// TIA Portal V20 export
// export: Created 2026-10-20T18:55:09.3234588Z, ExportSetting None, DisplayName Totally Integrated Automation Portal, DisplayVersion V20 Update 6, DisplayName TIA Portal Openness, DisplayVersion V20 Update 6, DisplayName TIA Portal Version Control Interface, DisplayVersion V20 Update 6, DisplayName SINAMICS Startdrive Advanced, DisplayVersion V20 SP1, DisplayName SINAMICS Startdrive G130, G150, S120, S150, SINAMICS MV, G220, S200, S210, DisplayVersion V20 SP1, DisplayName SINAMICS Startdrive G110M, G120, G120C, G120D, G120P, G115D, DisplayVersion V20 SP1, DisplayName STEP 7 Professional, DisplayVersion V20 Update 6, DisplayName STEP 7 Safety, DisplayVersion V20 Update 2, DisplayName WinCC Basic/Comfort/Advanced, DisplayVersion V20 Update 6, DisplayName WinCC Unified, DisplayVersion V20 Update 6
VAR_GLOBAL   // PLC tag table "IO_ET200_3"
   "C3204 - SENSOR CNV RIGHT (PALLET DETECT 1)" AT %I872.4 : Bool;
   "C3205 - SENSOR CNV RIGHT (PALLET DETECT 1)" AT %I874.4 : Bool;
   "C3207 - SENSOR CNV RIGHT (PALLET DETECT 1)" AT %I878.4 : Bool;
   "E-STOP L1 - CH1(3)" AT %I1662.0 : Bool;
   "E-STOP L2 - CH1(3)" AT %I1662.2 : Bool;
   "KEY REMOTE/LOCAL L1 - CH1(3)" AT %I1662.1 : Bool;
   "KEY REMOTE/LOCAL L2 - CH1(3)" AT %I1662.3 : Bool;
   "E-STOP L1 - CH2(3)" AT %I1662.4 : Bool;
   "KEY REMOTE/LOCAL L1 - CH2(3)" AT %I1662.5 : Bool;
   "E-STOP L2 - CH2(3)" AT %I1662.6 : Bool;
   "KEY REMOTE/LOCAL L2 - CH2(3)" AT %I1662.7 : Bool;
   "E-STOP L3 - CH1(3)" AT %I1670.0 : Bool;
   "KEY REMOTE/LOCAL L3 - CH1(3)" AT %I1670.1 : Bool;
   "E-STOP L4 - CH1(3)" AT %I1670.2 : Bool;
   "KEY REMOTE/LOCAL L4 - CH1(3)" AT %I1670.3 : Bool;
   "E-STOP L3 - CH2(3)" AT %I1670.4 : Bool;
   "KEY REMOTE/LOCAL L3 - CH2(3)" AT %I1670.5 : Bool;
   "E-STOP L4 - CH2(3)" AT %I1670.6 : Bool;
   "KEY REMOTE/LOCAL L4 - CH2(3)" AT %I1670.7 : Bool;
   "E-STOP L5 - CH1(3)" AT %I1678.0 : Bool;
   "KEY REMOTE/LOCAL L5 - CH1(3)" AT %I1678.1 : Bool;
   "E-STOP L6 - CH1(3)" AT %I1678.2 : Bool;
   "KEY REMOTE/LOCAL L6 - CH1(3)" AT %I1678.3 : Bool;
   "E-STOP L5 - CH2(3)" AT %I1678.4 : Bool;
   "KEY REMOTE/LOCAL L5 - CH2(3)" AT %I1678.5 : Bool;
   "E-STOP L6 - CH2(3)" AT %I1678.6 : Bool;
   "KEY REMOTE/LOCAL L6 - CH2(3)" AT %I1678.7 : Bool;
   "E-STOP L8 - CH1(3)" AT %I1686.2 : Bool;
   "KEY REMOTE/LOCAL L8 - CH1(3)" AT %I1686.3 : Bool;
   "E-STOP L8 - CH2(3)" AT %I1686.6 : Bool;
   "KEY REMOTE/LOCAL L8 - CH2(3)" AT %I1686.7 : Bool;
   "C3201 - SENSOR CNV RIGHT (PALLET DETECT 1)" AT %I866.4 : Bool;
   "C3201 - SHUTTLE IN POSITION 2" AT %I867.6 : Bool;
   "CVTD3 SENSOR CONVEYOR LEFT (PALLET DETECT 1)" AT %I140.2 : Bool;
   "C3201 - SENSOR CNV RIGHT (PALLET DETECT 2)" AT %I867.1 : Bool;
   "VTD3 DOCKING PINS EXTENDED 1" AT %I141.0 : Bool;
   "VTD3 LEVEL DETECT 1" AT %I141.7 : Bool;
   "C3201 - SENSOR CNV LEFT (FWD)" AT %I867.4 : Bool;
   "VTD3 DOCKING PINS EXTENDED 2" AT %I141.2 : Bool;
   "VTD3 LEVEL DETECT 2" AT %I141.6 : Bool;
   "C3201 - SHUTTLE IN POSITION 1" AT %I867.7 : Bool;
   "VTD3 DOCKING PINS RETRACTED 1" AT %I141.1 : Bool;
   "CVTD3 SENSOR CONVEYOR CENTER" AT %I140.3 : Bool;
   "VTD3 ULTIMATE SLOWDOWN" AT %I141.4 : Bool;
   "VTD3 ULTIMATE CREEP" AT %I141.5 : Bool;
   "CVTD3 SENSOR CONVEYOR RIGHT (PALLET DETECT 1)" AT %I140.5 : Bool;
   "CVTD3 SENSOR CONVEYOR LEFT (FWD)" AT %I140.1 : Bool;
   "VTD3 DOCKING PINS RETRACTED 2" AT %I141.3 : Bool;
   "C3201 - SENSOR CNV RIGHT (BWD)" AT %I866.5 : Bool;
   "C3201 - SENSOR CNV LEFT (PALLET DETECT 2)" AT %I867.0 : Bool;
   "C3201 - SENSOR CNV LEFT (PALLET DETECT 1)" AT %I867.5 : Bool;
   "CVTD3 SENSOR CONVEYOR RIGHT (BWD)" AT %I140.4 : Bool;
   "C3106 - SENSOR CNV RIGHT (PALLET DETECT 1)" AT %I861.5 : Bool;
   "C3208 - SENSOR CNV LEFT (FWD)" AT %I881.4 : Bool;
   "C3108 - SENSOR CNV LEFT (FWD)" AT %I864.5 : Bool;
   "C3107 - SENSOR CNV LEFT (PALLET DETECT 1)" AT %I862.4 : Bool;
   "C3107 - SENSOR CNV RIGHT (PALLET DETECT 2)" AT %I863.0 : Bool;
   "C3107 - SENSOR SAFETY PIN1 DOWN" AT %I863.3 : Bool;
   "C3208 - SENSOR SAFETY PIN1 UP" AT %I881.2 : Bool;
   "C3208 - SENSOR SAFETY PIN1 DOWN" AT %I881.3 : Bool;
   "C3108 - SENSOR SAFETY PIN1 DOWN" AT %I865.3 : Bool;
   "C3108 - SENSOR CNV RIGHT (PALLET DETECT 1)" AT %I865.5 : Bool;
   "C3207 - SENSOR CNV LEFT (PALLET DETECT 1)" AT %I879.1 : Bool;
   "C3106 - SENSOR SAFETY PIN1 DOWN" AT %I861.3 : Bool;
   "C3207 - SENSOR CNV RIGHT (PALLET DETECT 2)" AT %I879.5 : Bool;
   "C3106 - SENSOR CNV LEFT (PALLET DETECT 1)" AT %I860.4 : Bool;
   "C3108 - SENSOR CNV RIGHT (PALLET DETECT 2)" AT %I865.0 : Bool;
   "C3106 - SENSOR CNV LEFT (FWD)" AT %I860.5 : Bool;
   "C3206 - SENSOR CNV LEFT (PALLET DETECT 2)" AT %I877.0 : Bool;
   "C3207 - SENSOR CNV LEFT (FWD)" AT %I879.0 : Bool;
   "C3208 - SENSOR CNV RIGHT (PALLET DETECT 1)" AT %I880.4 : Bool;
   "C3208 - SENSOR CNV LEFT (PALLET DETECT 2)" AT %I881.0 : Bool;
   "C3106 - SENSOR CNV LEFT (PALLET DETECT 2)" AT %I861.1 : Bool;
   "C3108 - SENSOR CNV RIGHT (BWD)" AT %I865.4 : Bool;
   "C3206 - SENSOR CNV LEFT (FWD)" AT %I877.4 : Bool;
   "C3107 - SENSOR CNV RIGHT (BWD)" AT %I863.4 : Bool;
   "C3106 - SENSOR CNV RIGHT (BWD)" AT %I861.4 : Bool;
   "C3207 - SENSOR SAFETY PIN1 DOWN" AT %I879.3 : Bool;
   "C3108 - SENSOR CNV LEFT (PALLET DETECT 1)" AT %I864.4 : Bool;
   "C3108 - SHUTTLE IN POSITION 2" AT %I865.6 : Bool;
   "C3107 - SENSOR CNV LEFT (PALLET DETECT 2)" AT %I863.1 : Bool;
   "C3107 - SENSOR SAFETY PIN1 UP" AT %I863.2 : Bool;
   "C3106 - SHUTTLE IN POSITION 1" AT %I861.7 : Bool;
   "C3208 - SENSOR CNV LEFT (PALLET DETECT 1)" AT %I881.5 : Bool;
   "C3207 - SHUTTLE IN POSITION 1" AT %I879.7 : Bool;
   "C3208 - SENSOR CNV RIGHT (BWD)" AT %I880.5 : Bool;
   "C3108 - SENSOR SAFETY PIN1 UP" AT %I865.2 : Bool;
   "C3107 - SENSOR CNV RIGHT (PALLET DETECT 1)" AT %I863.5 : Bool;
   "C3207 - SENSOR CNV LEFT (PALLET DETECT 2)" AT %I879.4 : Bool;
   "C3207 - SENSOR CNV RIGHT (BWD)" AT %I878.5 : Bool;
   "C3207 - SENSOR SAFETY PIN1 UP" AT %I879.2 : Bool;
   "C3108 - SHUTTLE IN POSITION 1" AT %I865.7 : Bool;
   "C3106 - SENSOR CNV RIGHT (PALLET DETECT 2)" AT %I861.0 : Bool;
   "C3208 - SHUTTLE IN POSITION 1" AT %I881.7 : Bool;
   "C3106 - SHUTTLE IN POSITION 2" AT %I861.6 : Bool;
   "C3106 - SENSOR SAFETY PIN1 UP" AT %I861.2 : Bool;
   "C3206 - SENSOR CNV LEFT (PALLET DETECT 1)" AT %I877.5 : Bool;
   "C3107 - SENSOR CNV LEFT (FWD)" AT %I862.5 : Bool;
   "C3208 - SHUTTLE IN POSITION 2" AT %I881.6 : Bool;
   "C3206 - SENSOR CNV RIGHT (PALLET DETECT 2)" AT %I877.1 : Bool;
   "C3108 - SENSOR CNV LEFT (PALLET DETECT 2)" AT %I865.1 : Bool;
   "C3107 - SHUTTLE IN POSITION 2" AT %I863.6 : Bool;
   "C3208 - SENSOR CNV RIGHT (PALLET DETECT 2)" AT %I881.1 : Bool;
   "C3107 - SHUTTLE IN POSITION 1" AT %I863.7 : Bool;
   "C3207 - SHUTTLE IN POSITION 2" AT %I879.6 : Bool;
   "C3105 - SENSOR CNV LEFT (FWD)" AT %I858.5 : Bool;
   "C3104 - SENSOR CNV LEFT (PALLET DETECT 2)" AT %I857.1 : Bool;
   "C3104 - SENSOR CNV LEFT (FWD)" AT %I856.5 : Bool;
   "C3206 - SENSOR CNV RIGHT (PALLET DETECT 1)" AT %I876.0 : Bool;
   "C3104 - SHUTTLE IN POSITION 1" AT %I857.7 : Bool;
   "C3105 - SHUTTLE IN POSITION 1" AT %I859.7 : Bool;
   "C3205 - SENSOR CNV LEFT (FWD)" AT %I875.4 : Bool;
   "C3105 - SENSOR CNV LEFT (PALLET DETECT 1)" AT %I858.4 : Bool;
   "C3205 - SENSOR SAFETY PIN1 DOWN" AT %I875.3 : Bool;
   "C3105 - SHUTTLE IN POSITION 2" AT %I859.6 : Bool;
   "C3105 - SENSOR SAFETY PIN1 DOWN" AT %I859.3 : Bool;
   "C3206 - SENSOR CNV RIGHT (BWD)" AT %I876.1 : Bool;
   "C3206 - SENSOR SAFETY PIN1 DOWN" AT %I877.3 : Bool;
   "C3104 - SHUTTLE IN POSITION 2" AT %I857.6 : Bool;
   "C3206 - SENSOR SAFETY PIN1 UP" AT %I877.2 : Bool;
   "C3104 - SENSOR SAFETY PIN1 UP" AT %I857.2 : Bool;
   "C3104 - SENSOR CNV RIGHT (PALLET DETECT 2)" AT %I857.0 : Bool;
   "C3205 - SENSOR SAFETY PIN1 UP" AT %I875.2 : Bool;
   "C3105 - SENSOR CNV LEFT (PALLET DETECT 2)" AT %I859.1 : Bool;
   "C3205 - SENSOR CNV LEFT (PALLET DETECT 2)" AT %I875.0 : Bool;
   "C3105 - SENSOR CNV RIGHT (PALLET DETECT 1)" AT %I859.5 : Bool;
   "C3206 - SHUTTLE IN POSITION 1" AT %I877.7 : Bool;
   "C3104 - SENSOR CNV RIGHT (BWD)" AT %I857.4 : Bool;
   "C3205 - SENSOR CNV RIGHT (PALLET DETECT 2)" AT %I875.1 : Bool;
   "C3104 - SENSOR CNV RIGHT (PALLET DETECT 1)" AT %I857.5 : Bool;
   "C3205 - SHUTTLE IN POSITION 2" AT %I875.6 : Bool;
   "C3206 - SHUTTLE IN POSITION 2" AT %I877.6 : Bool;
   "C3105 - SENSOR CNV RIGHT (PALLET DETECT 2)" AT %I859.0 : Bool;
   "C3105 - SENSOR CNV RIGHT (BWD)" AT %I859.4 : Bool;
   "C3205 - SENSOR CNV RIGHT (BWD)" AT %I874.5 : Bool;
   "C3205 - SHUTTLE IN POSITION 1" AT %I875.7 : Bool;
   "C3104 - SENSOR SAFETY PIN1 DOWN" AT %I857.3 : Bool;
   "C3104 - SENSOR CNV LEFT (PALLET DETECT 1)" AT %I856.4 : Bool;
   "C3205 - SENSOR CNV LEFT (PALLET DETECT 1)" AT %I875.5 : Bool;
   "C3105 - SENSOR SAFETY PIN1 UP" AT %I859.2 : Bool;
   "C3204 - SENSOR CNV LEFT (PALLET DETECT 1)" AT %I873.5 : Bool;
   "C3102 - SENSOR CNV LEFT (PALLET DETECT 1)" AT %I536.4 : Bool;
   "C3102 - SENSOR SAFETY PIN1 DOWN" AT %I537.3 : Bool;
   "C3202 - SENSOR CNV LEFT (FWD)" AT %I869.4 : Bool;
   "C3204 - SENSOR CNV LEFT (PALLET DETECT 2)" AT %I873.0 : Bool;
   "C3203 - SENSOR CNV RIGHT (BWD)" AT %I870.5 : Bool;
   "C3203 - SENSOR CNV LEFT (FWD)" AT %I871.4 : Bool;
   "C3202 - SENSOR SAFETY PIN1 UP" AT %I869.2 : Bool;
   "C3204 - SENSOR SAFETY PIN1 DOWN" AT %I873.3 : Bool;
   "C3203 - SHUTTLE IN POSITION 1" AT %I871.7 : Bool;
   "C3102 - SENSOR CNV LEFT (FWD)" AT %I536.5 : Bool;
   "C3202 - SENSOR CNV LEFT (PALLET DETECT 1)" AT %I869.5 : Bool;
   "C3203 - SHUTTLE IN POSITION 2" AT %I871.6 : Bool;
   "C3202 - SHUTTLE IN POSITION 1" AT %I869.7 : Bool;
   "C3204 - SENSOR SAFETY PIN1 UP" AT %I873.2 : Bool;
   "C3203 - SENSOR CNV LEFT (PALLET DETECT 1)" AT %I871.5 : Bool;
   "C3102 - SENSOR CNV RIGHT (BWD)" AT %I537.4 : Bool;
   "C3203 - SENSOR CNV LEFT (PALLET DETECT 2)" AT %I871.0 : Bool;
   "C3102 - SHUTTLE IN POSITION 1" AT %I537.7 : Bool;
   "C3204 - SENSOR CNV LEFT (FWD)" AT %I873.4 : Bool;
   "C3202 - SENSOR CNV LEFT (PALLET DETECT 2)" AT %I869.0 : Bool;
   "C3204 - SHUTTLE IN POSITION 2" AT %I873.6 : Bool;
   "C3203 - SENSOR CNV RIGHT (PALLET DETECT 2)" AT %I871.1 : Bool;
   "C3202 - SENSOR CNV RIGHT (PALLET DETECT 1)" AT %I868.4 : Bool;
   "C3204 - SHUTTLE IN POSITION 1" AT %I873.7 : Bool;
   "C3204 - SENSOR CNV RIGHT (PALLET DETECT 2)" AT %I873.1 : Bool;
   "C3202 - SENSOR CNV RIGHT (BWD)" AT %I868.5 : Bool;
   "C3202 - SENSOR CNV RIGHT (PALLET DETECT 2)" AT %I869.1 : Bool;
   "C3102 - SENSOR SAFETY PIN1 UP" AT %I537.2 : Bool;
   "C3102 - SHUTTLE IN POSITION 2" AT %I537.6 : Bool;
   "C3203 - SENSOR SAFETY PIN1 DOWN" AT %I871.3 : Bool;
   "C3202 - SHUTTLE IN POSITION 2" AT %I869.6 : Bool;
   "C3102 - SENSOR CNV RIGHT (PALLET DETECT 1)" AT %I537.5 : Bool;
   "C3102 - SENSOR CNV LEFT (PALLET DETECT 2)" AT %I537.1 : Bool;
   "C3203 - SENSOR CNV RIGHT (PALLET DETECT 1)" AT %I870.4 : Bool;
   "C3202 - SENSOR SAFETY PIN1 DOWN" AT %I869.3 : Bool;
   "C3203 - SENSOR SAFETY PIN1 UP" AT %I871.2 : Bool;
   "C3102 - SENSOR CNV RIGHT (PALLET DETECT 2)" AT %I537.0 : Bool;
   "C3204 - SENSOR CNV RIGHT (BWD)" AT %I872.5 : Bool;
   "KEY REMOTE/LOCAL L7 - CH1(3)" AT %I1686.0 : Bool;
   "E-STOP L7 - CH1(3)" AT %I1686.1 : Bool;
   "KEY REMOTE/LOCAL L7 - CH2(3)" AT %I1686.4 : Bool;
   "E-STOP L7 - CH2(3)" AT %I1686.5 : Bool;
   "C3101 - SENSOR CNV RIGHT (PALLET DETECT 2)" AT %I498.4 : Bool;
   "C3101 - SHUTTLE IN POSITION 2" AT %I499.2 : Bool;
   "C3101 - SENSOR CNV LEFT (PALLET DETECT 2)" AT %I498.5 : Bool;
   "C3101 - SENSOR CNV LEFT (FWD)" AT %I498.3 : Bool;
   "C3101 - SENSOR CNV RIGHT (BWD)" AT %I498.0 : Bool;
   "C3101 - SENSOR CNV RIGHT (PALLET DETECT 1)" AT %I498.1 : Bool;
   "C3101 - SENSOR CNV LEFT (PALLET DETECT 1)" AT %I498.2 : Bool;
   "C3101 - SHUTTLE IN POSITION 1" AT %I499.3 : Bool;
   "C3103 - SENSOR SAFETY PIN1 DOWN" AT %I539.1 : Bool;
   "C3103 - SHUTTLE IN POSITION 2" AT %I538.6 : Bool;
   "C3103 - SENSOR CNV RIGHT (PALLET DETECT 2)" AT %I538.4 : Bool;
   "C3103 - SENSOR SAFETY PIN1 UP" AT %I539.0 : Bool;
   "C3103 - SENSOR CNV RIGHT (BWD)" AT %I538.0 : Bool;
   "C3103 - SENSOR CNV LEFT (PALLET DETECT 2)" AT %I538.5 : Bool;
   "C3103 - SENSOR CNV RIGHT (PALLET DETECT 1)" AT %I538.1 : Bool;
   "C3103 - SENSOR CNV LEFT (FWD)" AT %I538.3 : Bool;
   "C3103 - SHUTTLE IN POSITION 1" AT %I538.7 : Bool;
   "C3103 - SENSOR CNV LEFT (PALLET DETECT 1)" AT %I538.2 : Bool;
   "CVTD3 OVERHANG RIGHT" AT %I140.6 : Bool;
   "CVTD3 OVERHANG LEFT" AT %I140.7 : Bool;
END_VAR
